FUNCTION_BLOCK PvPorcentagem (* Pv em porcentagem da faixa de medicao (PvMin..PvMax), calculado no CLP para a IHM *)
  (* Standard: 61499-2 *)
  (* Version 1.0, 06/11/2026, Hidryco, Hidryco, 1.0: PvPct = (Pv - PvMin) / (PvMax - PvMin) x 100; faixa nula = 0. Sem limitar a 0..100 (acima da faixa aparece acima de 100). *)
  PACKAGE SE.Nereda;
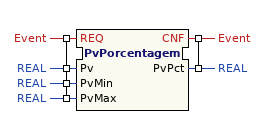
  EVENT_INPUT
    REQ WITH Pv, PvMin, PvMax; (* Novo valor medido *)
  END_EVENT
  EVENT_OUTPUT
    CNF WITH PvPct; (* Porcentagem atualizada *)
  END_EVENT
  VAR_INPUT
    Pv : REAL; (* Valor medido (unidade de engenharia) *)
    PvMin : REAL; (* Inicio da faixa (4 mA) *)
    PvMax : REAL; (* Fim da faixa (20 mA) *)
  END_VAR
  VAR_OUTPUT
    PvPct : REAL; (* Valor em porcentagem da faixa *)
  END_VAR
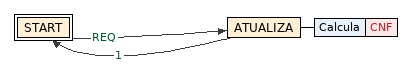
  EC_STATES
    START; (* Estado inicial *)
    ATUALIZA : Calcula -> CNF; (* Calcula e emite *)
  END_STATES
  EC_TRANSITIONS
    START TO ATUALIZA := REQ;
    ATUALIZA TO START := 1;
  END_TRANSITIONS
  ALGORITHM Calcula IN ST: (* Porcentagem da faixa *)
IF PvMax <> PvMin THEN
    PvPct := (Pv - PvMin) / (PvMax - PvMin) * 100.0;
ELSE
    PvPct := 0.0;
END_IF;
  END_ALGORITHM
END_FUNCTION_BLOCK
